(* IEC 61131-3 sources: PLC-Static-Analysis/modules/plc-rules/src/test/resources/PLCA-L022, 2 files *)

(* ---- compliant.st ---- *)
PROGRAM P_L022ok
VAR
    n : INT;
    m : INT;
    r : REAL;
    b : BOOL;
    c : BOOL;
    q : BOOL;
    aData : ARRAY[1..10] OF INT;
END_VAR
FOR n := 1 TO 10 DO
    IF aData[n] > 100 THEN
        m := n;
        EXIT;
    END_IF
END_FOR
WHILE TRUE DO
    IF NOT b THEN
        EXIT;
    END_IF
    m := m + 1;
    IF m > 5 THEN
        EXIT;
    END_IF
    q := TRUE;
    EXIT;
END_WHILE
FOR n := 1 TO 10 DO
    IF aData[n] = 0 THEN
        CONTINUE;
    END_IF
    m := n;
    EXIT;
END_FOR
END_PROGRAM

(* ---- noncompliant.st ---- *)
PROGRAM P_L022
VAR
    n : INT;
    m : INT;
    r : REAL;
    b : BOOL;
    c : BOOL;
    q : BOOL;
    aData : ARRAY[1..10] OF INT;
END_VAR
FOR n := 1 TO 10 DO // PLCA-L022
    IF aData[n] > 100 THEN
        m := n;
    END_IF
    EXIT;
END_FOR
WHILE b DO // PLCA-L022
    m := m + 1;
    RETURN;
END_WHILE
END_PROGRAM
